TYPE ST_Signals :
STRUCT
    {attribute 'TagName' := 'ID'}
    signal : STRING(255);
    
    {attribute 'FieldName' := 'Value'}
    value : LREAL := -1;
	
END_STRUCT
END_TYPE

(* stored: Version 1.1.0.1
   DUT ST_Signals: Id {95451f05-13c1-45b3-8a34-da3612fda24e} *)
